(* Logix 5000 project; controller R400_500_XLS vendor 1 type 14 code 216 rev 31.11; software revision 31.01; part 26 of 32 *)
(* tags used below, declared in another part *)
   Abort1 : DINT;   // Not Used
   Alarm : SINT;   // Wait 3 seconds
   AlarmAcked : BOOL;   // Alarm has been acked
   bAlrm : BOOL[64];
   Chem_Pump : UDT_CHEM_PUMP[4];   // Chemical Pump flow rate
   ChemPumpIndex : DINT;
   CycExcBuffer : UDT_CYCLE;
   CycleSequence : UDT_CYCLE_SEQUENCE;
   Delta_T : REAL;
   DRYING : DINT;   // Drying id number
   F1rinse : DINT;   // Not Used
   F2rinse : DINT;   // Not Used
   F3rinse : DINT;   // Not Used
   FC22_SumpWaterVolume : REAL;   // Water volume
   FC22_Tran1 : BOOL;   // First transition
   FC22_Tran3 : BOOL;   // Third transition
   FC22_Tran4 : BOOL;   // Fourth transition
   FC22_WashIndex : SINT;
   HeatSmp : DINT;
   HighLimt : REAL;
   I_Pw_Tnk_Lvl_Sw_Deb : BOOL;   // Debounced pure water tank level switch (100ms)
   Inj_Time : SINT;   // Time based chemical injection steps
   LowLimt : REAL;
   M : DINT[5];   // Memory Bits
   MaxPressRecord : REAL;
   MinPressRecord : REAL;
   Neutral : SINT;
   ONS_FC17_1 : BOOL;
   ONS_FC17_2 : BOOL;
   ONS_FC22 : SINT;
   ONS_FC40 : SINT;
   ONS_WSH30 : SINT;
   PrintPressureDelay : DINT;
   PumpLowFRinse : DINT;   // Delay for pump low speed during final rinse treatment
   PumpLowPW_W_R : DINT;   // Delay for pump low speed during pre-wash, wash and rinse treatments
   PURE_WATER_HEATING_TIME : DINT;   // Time before an alarm is thrown when the pure water tank is heating
   PureWaterTankFilling : BOOL;   // Start PWT filling
   PW_HeatSp_5 : REAL;
   PW_HeatSp_X : REAL;
   PWHeat : SINT;
   Run : DINT;
   Service : DINT[2];   // Unused Service Mode Memory Bit
   StartPump1 : BOOL;   // Pump Low Speed
   StartPump2 : BOOL;   // Pump High Speed
   StartPump3 : BOOL;   // Main Pump running
   SUMP_HIGH_VOLUME_400 : REAL;   // High sump volume
   SUMP_HIGH_VOLUME_500 : REAL;
   SUMP_LOW_VOLUME_400 : REAL;   // Low sump volume
   SUMP_LOW_VOLUME_500 : REAL;
   SumpWaterVolume : DINT;   // Sump Water Volume 0 =Low 1= High
   T0_Temp : REAL;
   T1_Temp : REAL;
   TempChange : BOOL;
   Tmr : TIMER[107];
   Trt_PrWsh : DINT;
   Trt_Rinse : DINT;   // Rinse steps
   Trt_Wsh : DINT;
   WASH_1 : DINT;   // Wash 1 id number
   WASH_5 : DINT;   // Wash 5 id number
   WSH56_StartPump : BOOL;   // Start pump signal
   bPureWaterFillingAuthorization : BOOL;   // Pure Water Filling Authorization Signal
   I_Chm_1_Lvl_Sw : BOOL;   // Chemical Pump #1 level switch
   I_Chm_2_Lvl_Sw : BOOL;   // Chemical Pump #2 level switch
   I_Chm_3_Lvl_Sw : BOOL;   // Chemical Pump #3 level switch
   I_Chm_4_Lvl_Sw : BOOL;   // Chemical Pump #4 level switch
   I_MCR : BOOL;   // MCR input
   I_Mtr_Ovrld : BOOL;   // Motor overload
   I_Shlf_Sw : BOOL;   // Shelf switch
   PmpPres : REAL;
   PureWaterTankDrainingDeadLeg : BOOL;
   PureWaterTankFillingRequest : BOOL;
   PureWaterTankTemp : REAL;   // Pure water tank temperature
   Q_Pw_Tnk_Stm_Vlve : BOOL;   // PWT Steam Valve / Electric Heater
   SPV_19 : BOOL;   // Screen 80 Enabled/Disabled Pump pressure monitoring
   tDelayBeforeTankFillingAuthAlarm : TIMER;
   Tpb : DINT[11];
   tPureWaterTankClosingDelay : TIMER;
   TreatmentPtr : DINT;
   Unit : Hrdwre;   // Unit Configuration
(* MainProgram, continued *)

ROUTINE WSH_27_WSH_28_PURE_WATER_TANK   (* ladder *)
// This routine manages the filling, the draining and the heating of the pure water tank
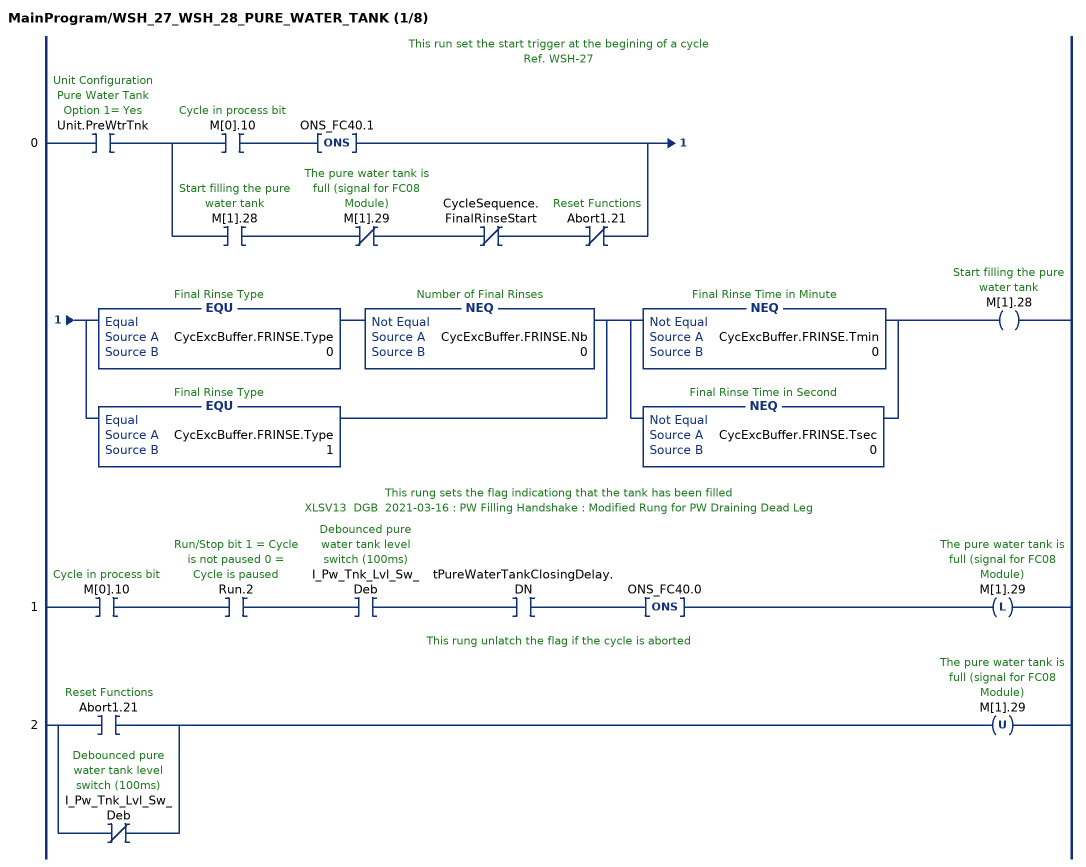
   // This run set the start trigger at the begining of a cycle
   // Ref. WSH-27
   0: XIC(Unit.PreWtrTnk)[XIC(M[0].10) ONS(ONS_FC40.1) ,XIC(M[1].28) XIO(M[1].29) XIO(CycleSequence.FinalRinseStart) XIO(Abort1.21) ][EQU(CycExcBuffer.FRINSE.Type,0) NEQ(CycExcBuffer.FRINSE.Nb,0) ,EQU(CycExcBuffer.FRINSE.Type,1) ][NEQ(CycExcBuffer.FRINSE.Tmin,0) ,NEQ(CycExcBuffer.FRINSE.Tsec,0) ]OTE(M[1].28);
   // This rung sets the flag indicationg that the tank has been filled
   // XLSV13  DGB  2021-03-16 : PW Filling Handshake : Modified Rung for PW Draining Dead Leg
   1: XIC(M[0].10)XIC(Run.2)XIC(I_Pw_Tnk_Lvl_Sw_Deb)XIC(tPureWaterTankClosingDelay.DN)ONS(ONS_FC40.0)OTL(M[1].29);
   // This rung unlatch the flag if the cycle is aborted
   2: [XIC(Abort1.21) ,XIO(I_Pw_Tnk_Lvl_Sw_Deb) ]OTU(M[1].29);
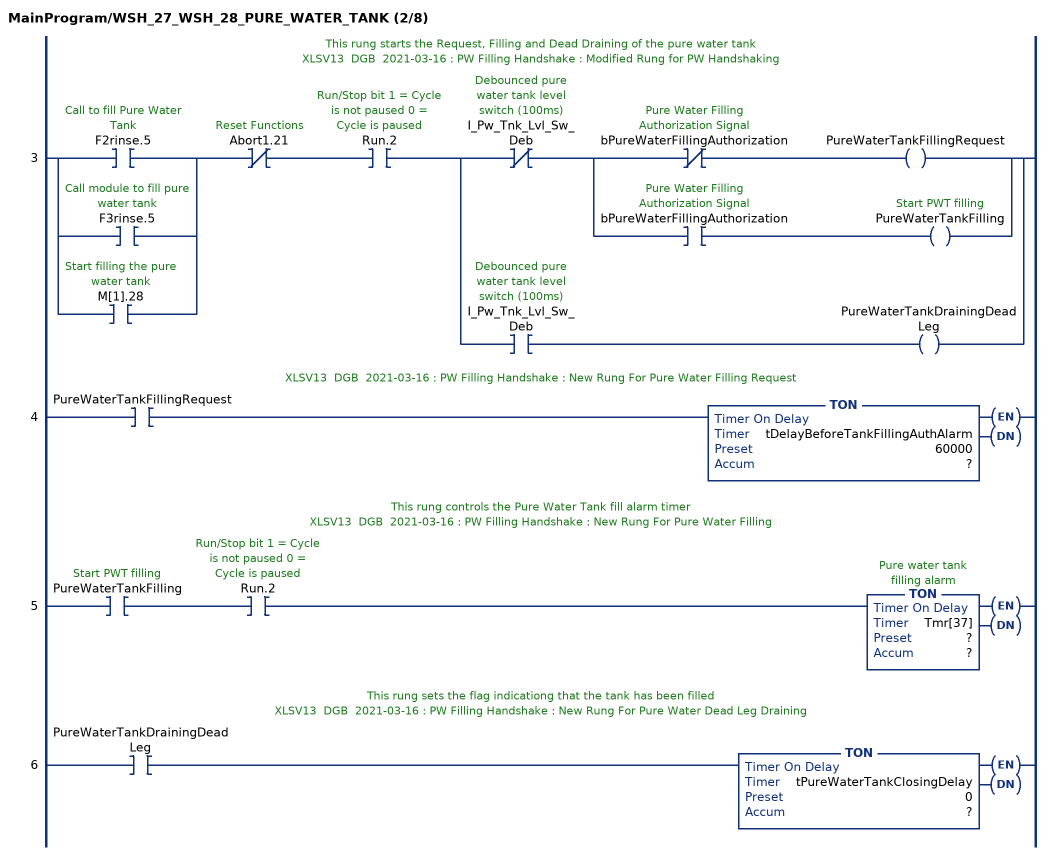
   // This rung starts the Request, Filling and Dead Draining of the pure water tank
   // XLSV13  DGB  2021-03-16 : PW Filling Handshake : Modified Rung for PW Handshaking
   3: [XIC(F2rinse.5) ,XIC(F3rinse.5) ,XIC(M[1].28) ]XIO(Abort1.21)XIC(Run.2)[XIO(I_Pw_Tnk_Lvl_Sw_Deb) [XIO(bPureWaterFillingAuthorization) OTE(PureWaterTankFillingRequest) ,XIC(bPureWaterFillingAuthorization) OTE(PureWaterTankFilling) ] ,XIC(I_Pw_Tnk_Lvl_Sw_Deb) OTE(PureWaterTankDrainingDeadLeg) ];
   // XLSV13  DGB  2021-03-16 : PW Filling Handshake : New Rung For Pure Water Filling Request
   4: XIC(PureWaterTankFillingRequest)TON(tDelayBeforeTankFillingAuthAlarm,?,?);
   // This rung controls the Pure Water Tank fill alarm timer
   // XLSV13  DGB  2021-03-16 : PW Filling Handshake : New Rung For Pure Water Filling
   5: XIC(PureWaterTankFilling)XIC(Run.2)TON(Tmr[37],?,?);
   // This rung sets the flag indicationg that the tank has been filled
   // XLSV13  DGB  2021-03-16 : PW Filling Handshake : New Rung For Pure Water Dead Leg Draining
   6: XIC(PureWaterTankDrainingDeadLeg)TON(tPureWaterTankClosingDelay,?,?);
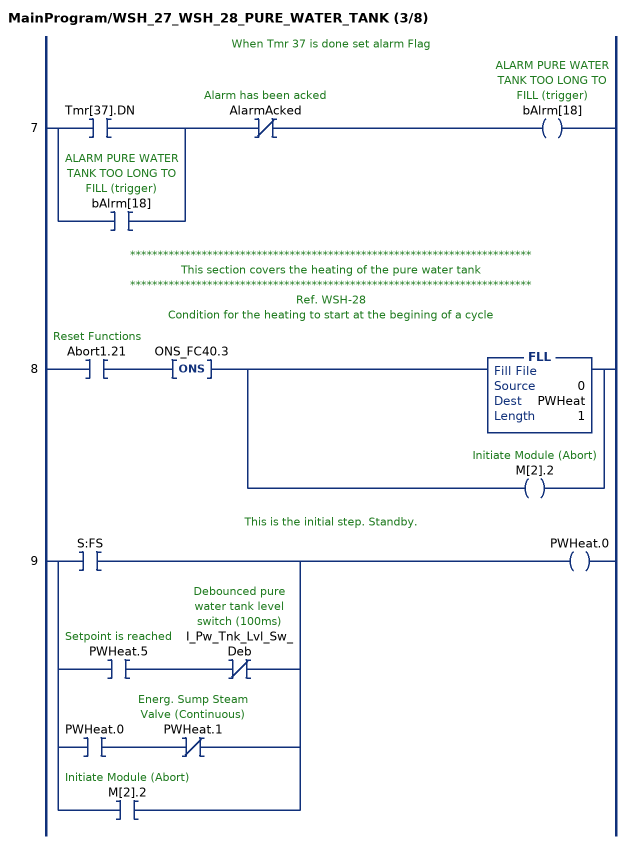
   // When Tmr 37 is done set alarm Flag
   7: [XIC(Tmr[37].DN) ,XIC(bAlrm[18]) ]XIO(AlarmAcked)OTE(bAlrm[18]);
   // *************************************************************************
   // This section covers the heating of the pure water tank
   // *************************************************************************
   // Ref. WSH-28
   // Condition for the heating to start at the begining of a cycle
   8: XIC(Abort1.21)ONS(ONS_FC40.3)[FLL(0,PWHeat,1) ,OTE(M[2].2) ];
   // This is the initial step. Standby.
   9: [XIC(S:FS) ,XIC(PWHeat.5) XIO(I_Pw_Tnk_Lvl_Sw_Deb) ,XIC(PWHeat.0) XIO(PWHeat.1) ,XIC(M[2].2) ]OTE(PWHeat.0);
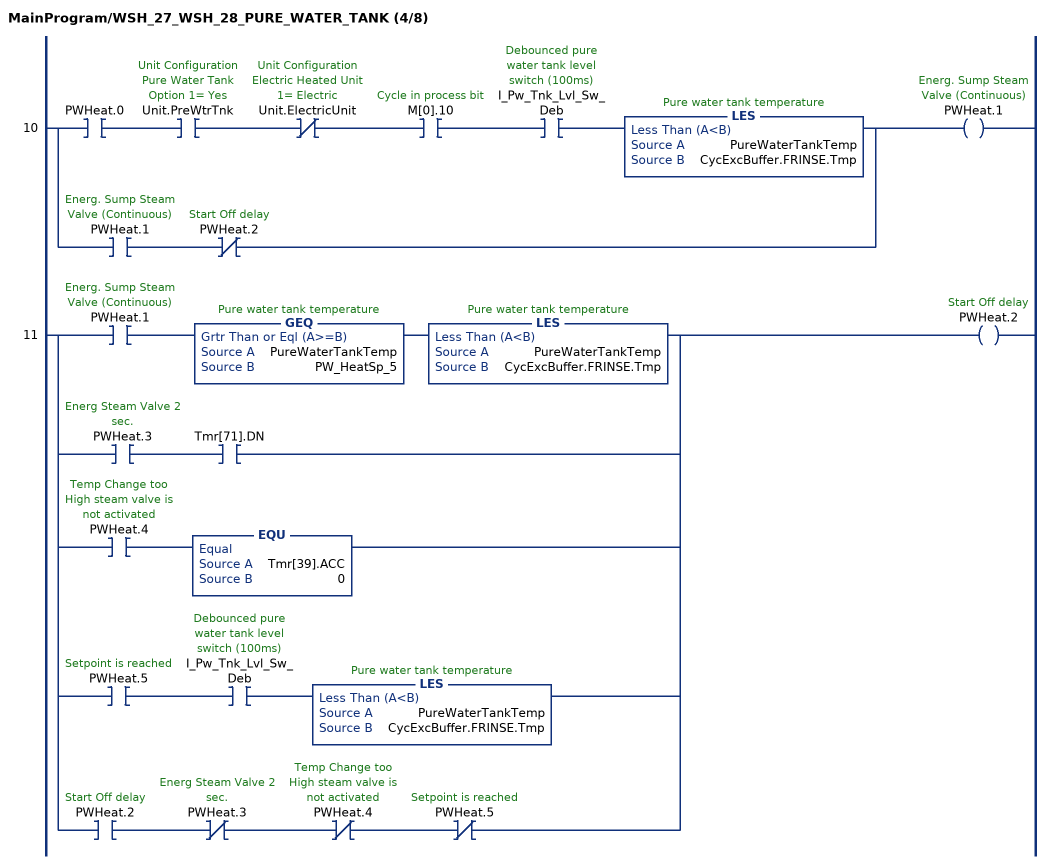
   10: [XIC(PWHeat.0) XIC(Unit.PreWtrTnk) XIO(Unit.ElectricUnit) XIC(M[0].10) XIC(I_Pw_Tnk_Lvl_Sw_Deb) LES(PureWaterTankTemp,CycExcBuffer.FRINSE.Tmp) ,XIC(PWHeat.1) XIO(PWHeat.2) ]OTE(PWHeat.1);
   11: [XIC(PWHeat.1) GEQ(PureWaterTankTemp,PW_HeatSp_5) LES(PureWaterTankTemp,CycExcBuffer.FRINSE.Tmp) ,XIC(PWHeat.3) XIC(Tmr[71].DN) ,XIC(PWHeat.4) EQU(Tmr[39].ACC,0) ,XIC(PWHeat.5) XIC(I_Pw_Tnk_Lvl_Sw_Deb) LES(PureWaterTankTemp,CycExcBuffer.FRINSE.Tmp) ,XIC(PWHeat.2) XIO(PWHeat.3) XIO(PWHeat.4) XIO(PWHeat.5) ]OTE(PWHeat.2);
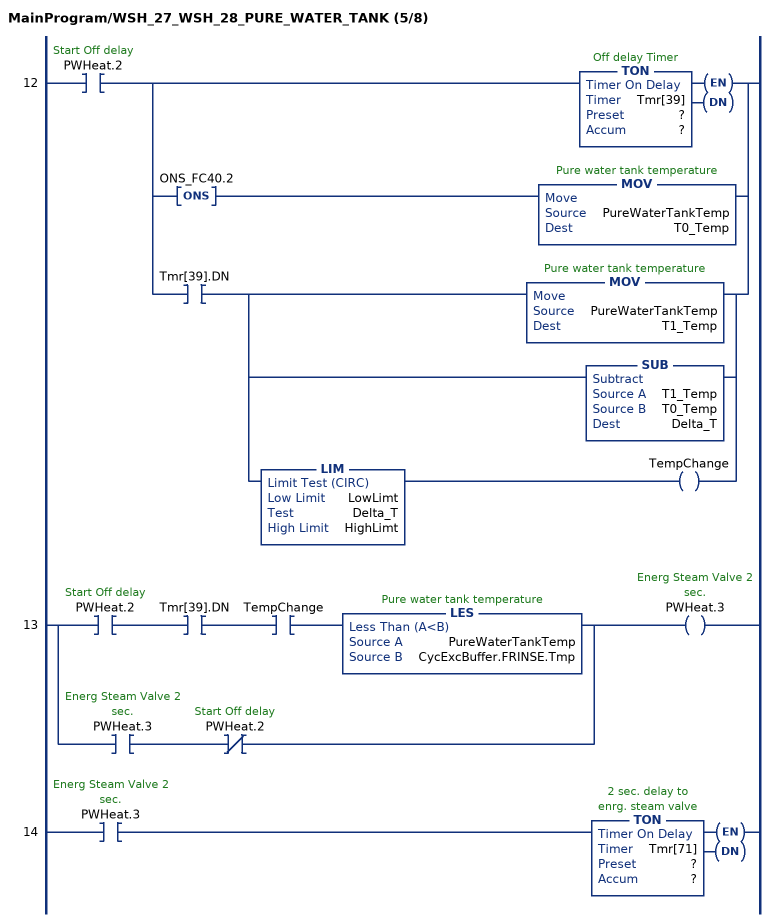
   12: XIC(PWHeat.2)[TON(Tmr[39],?,?) ,ONS(ONS_FC40.2) MOV(PureWaterTankTemp,T0_Temp) ,XIC(Tmr[39].DN) [MOV(PureWaterTankTemp,T1_Temp) ,SUB(T1_Temp,T0_Temp,Delta_T) ,LIM(LowLimt,Delta_T,HighLimt) OTE(TempChange) ] ];
   13: [XIC(PWHeat.2) XIC(Tmr[39].DN) XIC(TempChange) LES(PureWaterTankTemp,CycExcBuffer.FRINSE.Tmp) ,XIC(PWHeat.3) XIO(PWHeat.2) ]OTE(PWHeat.3);
   14: XIC(PWHeat.3)TON(Tmr[71],?,?);
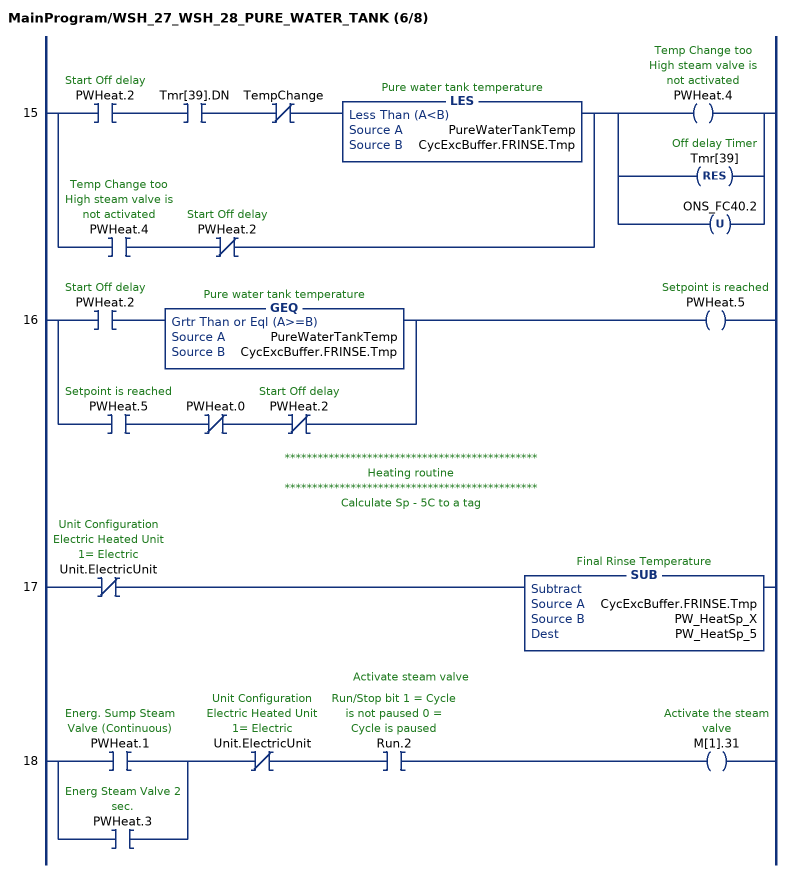
   15: [XIC(PWHeat.2) XIC(Tmr[39].DN) XIO(TempChange) LES(PureWaterTankTemp,CycExcBuffer.FRINSE.Tmp) ,XIC(PWHeat.4) XIO(PWHeat.2) ][OTE(PWHeat.4) ,RES(Tmr[39]) ,OTU(ONS_FC40.2) ];
   16: [XIC(PWHeat.2) GEQ(PureWaterTankTemp,CycExcBuffer.FRINSE.Tmp) ,XIC(PWHeat.5) XIO(PWHeat.0) XIO(PWHeat.2) ]OTE(PWHeat.5);
   // **********************************************
   // Heating routine
   // **********************************************
   // Calculate Sp - 5C to a tag
   17: XIO(Unit.ElectricUnit)SUB(CycExcBuffer.FRINSE.Tmp,PW_HeatSp_X,PW_HeatSp_5);
   // Activate steam valve
   18: [XIC(PWHeat.1) ,XIC(PWHeat.3) ]XIO(Unit.ElectricUnit)XIC(Run.2)OTE(M[1].31);
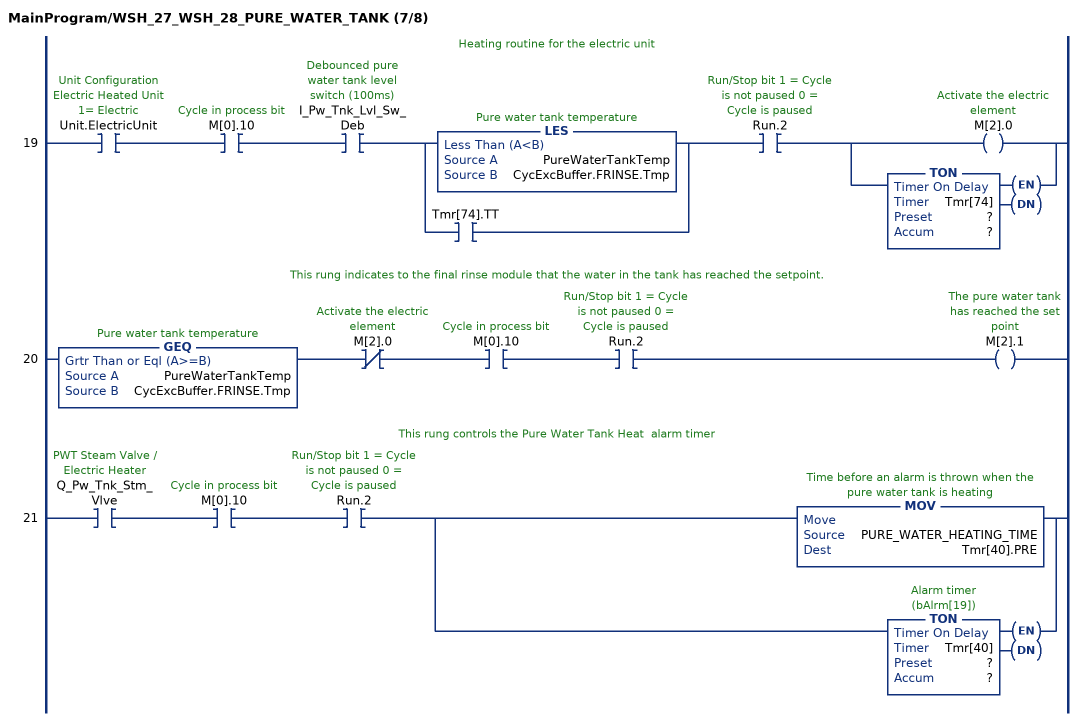
   // Heating routine for the electric unit
   19: XIC(Unit.ElectricUnit)XIC(M[0].10)XIC(I_Pw_Tnk_Lvl_Sw_Deb)[LES(PureWaterTankTemp,CycExcBuffer.FRINSE.Tmp) ,XIC(Tmr[74].TT) ]XIC(Run.2)[OTE(M[2].0) ,TON(Tmr[74],?,?) ];
   // This rung indicates to the final rinse module that the water in the tank has reached the setpoint.
   20: GEQ(PureWaterTankTemp,CycExcBuffer.FRINSE.Tmp)XIO(M[2].0)XIC(M[0].10)XIC(Run.2)OTE(M[2].1);
   // This rung controls the Pure Water Tank Heat  alarm timer
   21: XIC(Q_Pw_Tnk_Stm_Vlve)XIC(M[0].10)XIC(Run.2)[MOV(PURE_WATER_HEATING_TIME,Tmr[40].PRE) ,TON(Tmr[40],?,?) ];
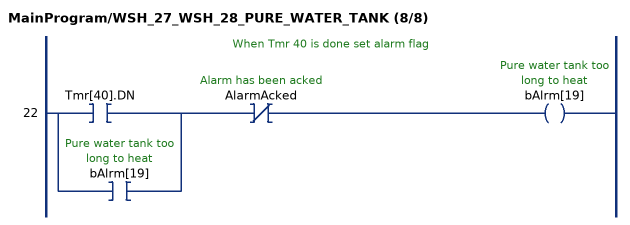
   // When Tmr 40 is done set alarm flag
   22: [XIC(Tmr[40].DN) ,XIC(bAlrm[19]) ]XIO(AlarmAcked)OTE(bAlrm[19]);
END_ROUTINE

ROUTINE WSH_29_START_PUMP   (* ladder *)
// This module starts the main pump
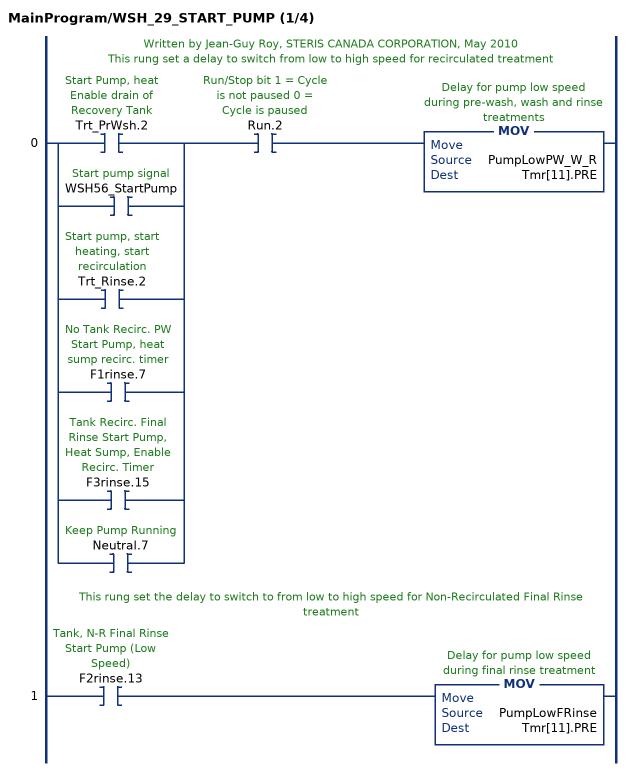
   // Written by Jean-Guy Roy, STERIS CANADA CORPORATION, May 2010
   // This rung set a delay to switch from low to high speed for recirculated treatment
   0: [XIC(Trt_PrWsh.2) ,XIC(WSH56_StartPump) ,XIC(Trt_Rinse.2) ,XIC(F1rinse.7) ,XIC(F3rinse.15) ,XIC(Neutral.7) ]XIC(Run.2)MOV(PumpLowPW_W_R,Tmr[11].PRE);
   // This rung set the delay to switch to from low to high speed for Non-Recirculated Final Rinse treatment
   1: XIC(F2rinse.13)MOV(PumpLowFRinse,Tmr[11].PRE);
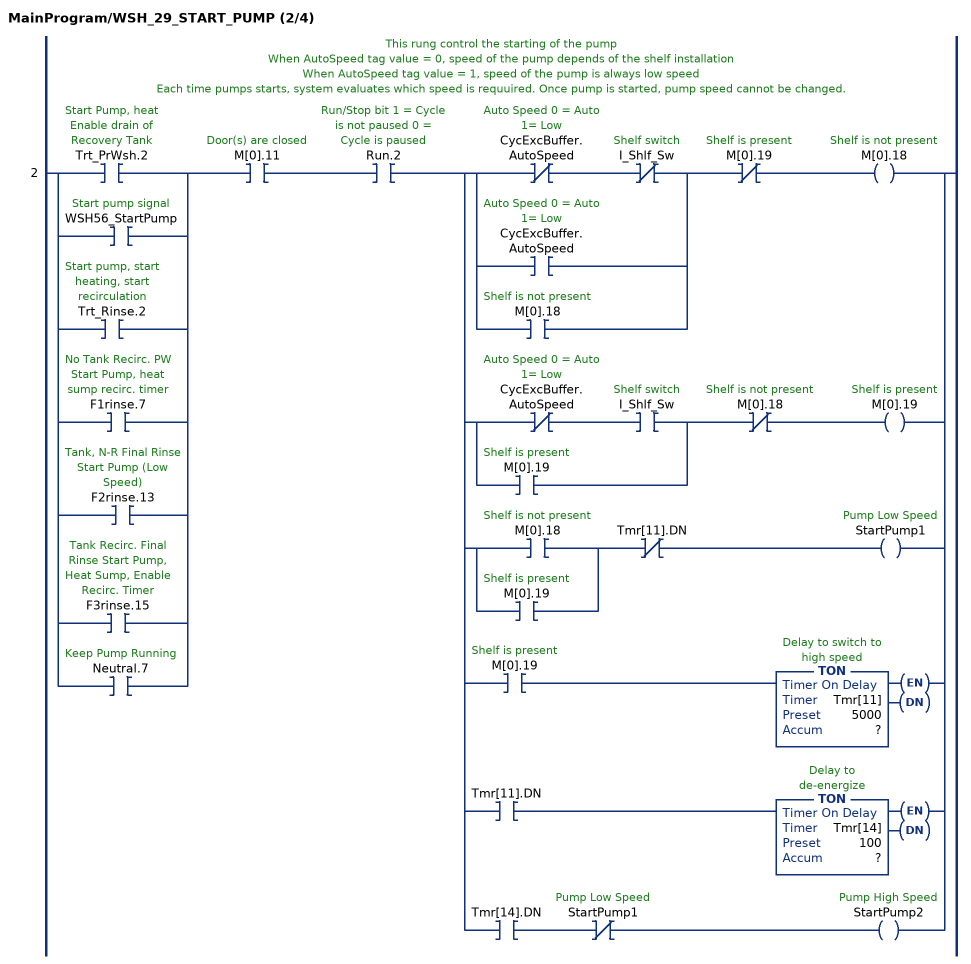
   // This rung control the starting of the pump
   // When AutoSpeed tag value = 0, speed of the pump depends of the shelf installation
   // When AutoSpeed tag value = 1, speed of the pump is always low speed
   // Each time pumps starts, system evaluates which speed is requuired. Once pump is started, pump speed cannot be changed.
   2: [XIC(Trt_PrWsh.2) ,XIC(WSH56_StartPump) ,XIC(Trt_Rinse.2) ,XIC(F1rinse.7) ,XIC(F2rinse.13) ,XIC(F3rinse.15) ,XIC(Neutral.7) ]XIC(M[0].11)XIC(Run.2)[[XIO(CycExcBuffer.AutoSpeed) XIO(I_Shlf_Sw) ,XIC(CycExcBuffer.AutoSpeed) ,XIC(M[0].18) ] XIO(M[0].19) OTE(M[0].18) ,[XIO(CycExcBuffer.AutoSpeed) XIC(I_Shlf_Sw) ,XIC(M[0].19) ] XIO(M[0].18) OTE(M[0].19) ,[XIC(M[0].18) ,XIC(M[0].19) ] XIO(Tmr[11].DN) OTE(StartPump1) ,XIC(M[0].19) TON(Tmr[11],?,?) ,XIC(Tmr[11].DN) TON(Tmr[14],?,?) ,XIC(Tmr[14].DN) XIO(StartPump1) OTE(StartPump2) ];
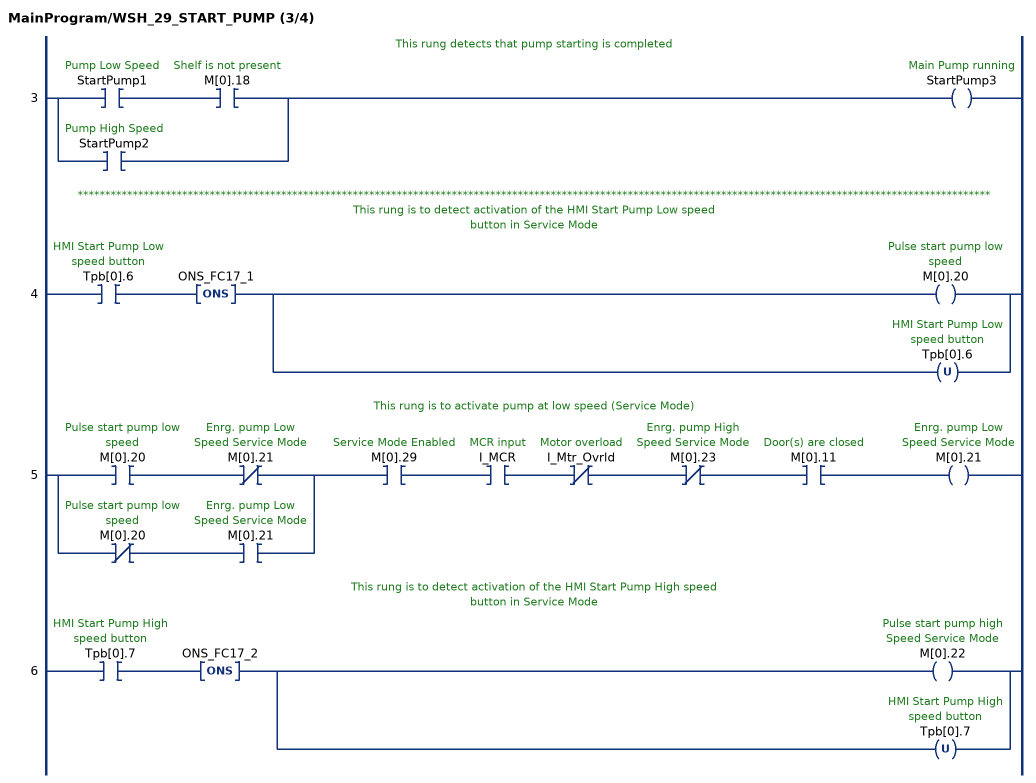
   // This rung detects that pump starting is completed
   3: [XIC(StartPump1) XIC(M[0].18) ,XIC(StartPump2) ]OTE(StartPump3);
   // **********************************************************************************************************************************************************************
   // This rung is to detect activation of the HMI Start Pump Low speed
   // button in Service Mode
   4: XIC(Tpb[0].6)ONS(ONS_FC17_1)[OTE(M[0].20) ,OTU(Tpb[0].6) ];
   // This rung is to activate pump at low speed (Service Mode)
   5: [XIC(M[0].20) XIO(M[0].21) ,XIO(M[0].20) XIC(M[0].21) ]XIC(M[0].29)XIC(I_MCR)XIO(I_Mtr_Ovrld)XIO(M[0].23)XIC(M[0].11)OTE(M[0].21);
   // This rung is to detect activation of the HMI Start Pump High speed
   // button in Service Mode
   6: XIC(Tpb[0].7)ONS(ONS_FC17_2)[OTE(M[0].22) ,OTU(Tpb[0].7) ];
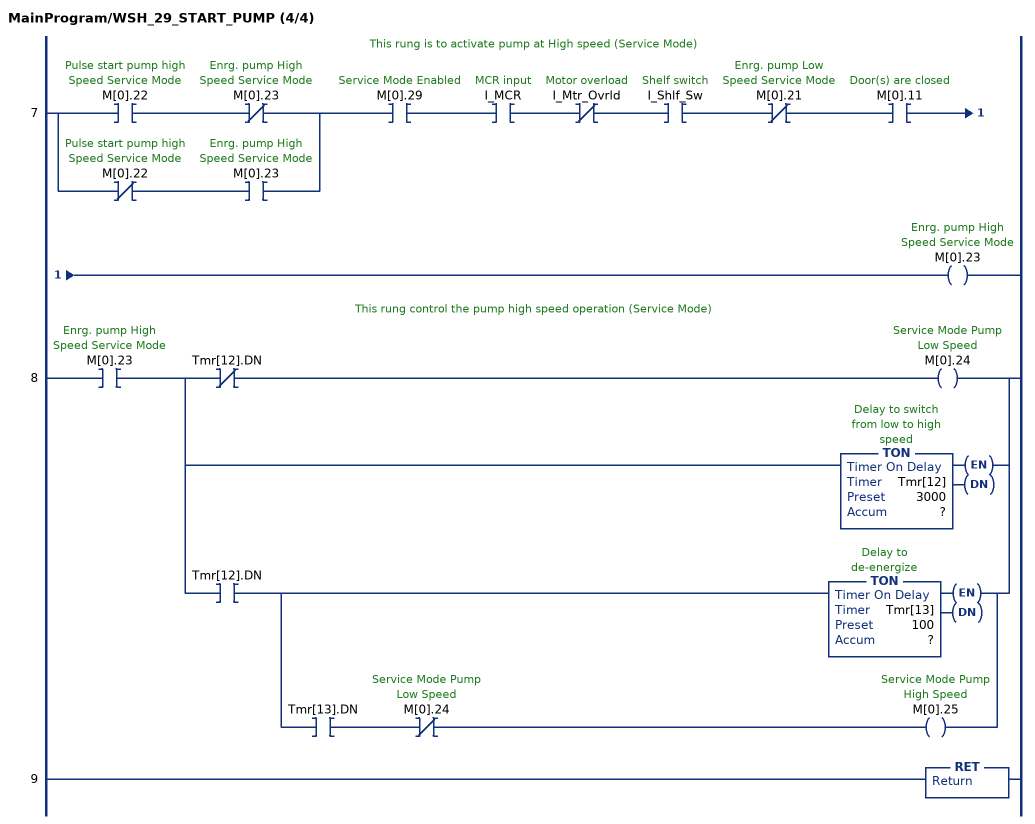
   // This rung is to activate pump at High speed (Service Mode)
   7: [XIC(M[0].22) XIO(M[0].23) ,XIO(M[0].22) XIC(M[0].23) ]XIC(M[0].29)XIC(I_MCR)XIO(I_Mtr_Ovrld)XIC(I_Shlf_Sw)XIO(M[0].21)XIC(M[0].11)OTE(M[0].23);
   // This rung control the pump high speed operation (Service Mode)
   8: XIC(M[0].23)[XIO(Tmr[12].DN) OTE(M[0].24) ,TON(Tmr[12],?,?) ,XIC(Tmr[12].DN) [TON(Tmr[13],?,?) ,XIC(Tmr[13].DN) XIO(M[0].24) OTE(M[0].25) ] ];
   9: RET();
END_ROUTINE

ROUTINE WSH_30_MONITOR_PRESSURE   (* ladder *)
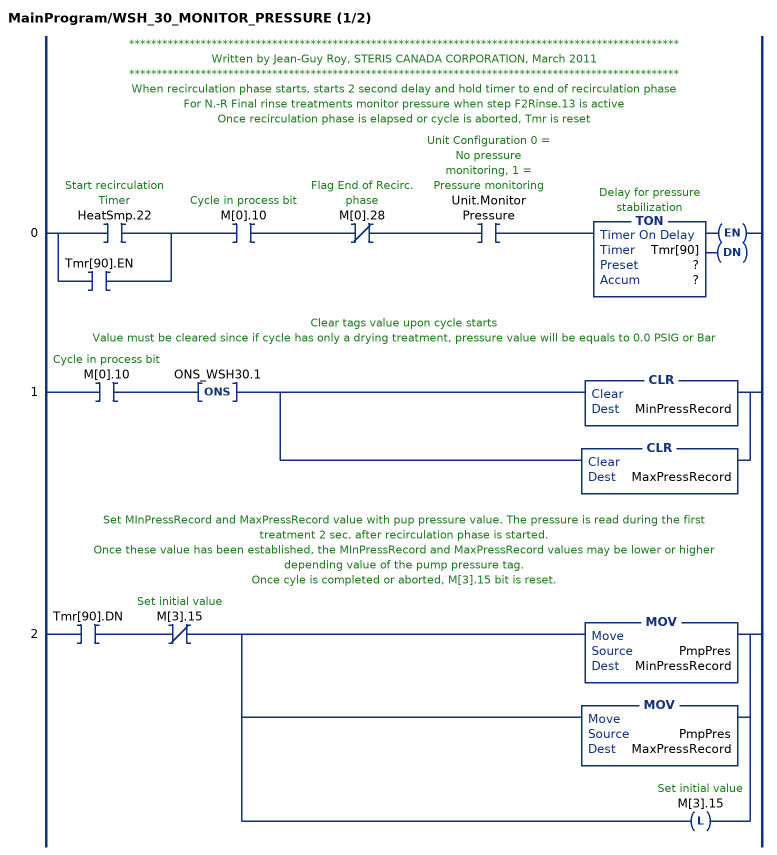
   // ****************************************************************************************************
   // Written by Jean-Guy Roy, STERIS CANADA CORPORATION, March 2011
   // ****************************************************************************************************
   // When recirculation phase starts, starts 2 second delay and hold timer to end of recirculation phase
   // For N.-R Final rinse treatments monitor pressure when step F2Rinse.13 is active
   // Once recirculation phase is elapsed or cycle is aborted, Tmr is reset
   0: [XIC(HeatSmp.22) ,XIC(Tmr[90].EN) ]XIC(M[0].10)XIO(M[0].28)XIC(Unit.MonitorPressure)TON(Tmr[90],?,?);
   // Clear tags value upon cycle starts
   // Value must be cleared since if cycle has only a drying treatment, pressure value will be equals to 0.0 PSIG or Bar
   1: XIC(M[0].10)ONS(ONS_WSH30.1)[CLR(MinPressRecord) ,CLR(MaxPressRecord) ];
   // Set MInPressRecord and MaxPressRecord value with pup pressure value. The pressure is read during the first treatment 2 sec. after recirculation phase is started.
   // Once these value has been established, the MInPressRecord and MaxPressRecord values may be lower or higher depending value of the pump pressure tag.
   // Once cyle is completed or aborted, M[3].15 bit is reset.
   2: XIC(Tmr[90].DN)XIO(M[3].15)[MOV(PmpPres,MinPressRecord) ,MOV(PmpPres,MaxPressRecord) ,OTL(M[3].15) ];
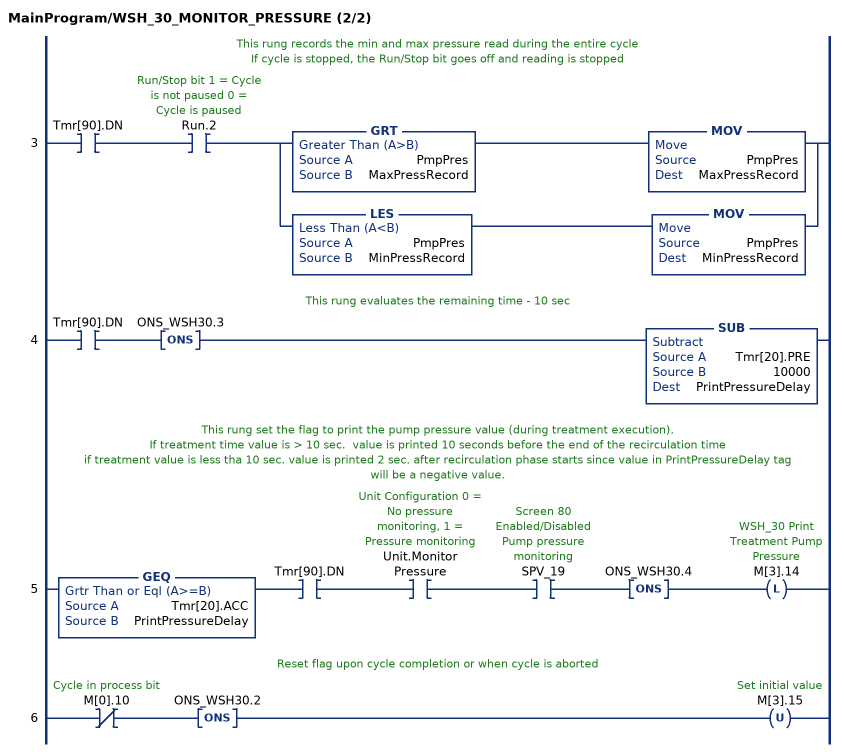
   // This rung records the min and max pressure read during the entire cycle
   // If cycle is stopped, the Run/Stop bit goes off and reading is stopped
   3: XIC(Tmr[90].DN)XIC(Run.2)[GRT(PmpPres,MaxPressRecord) MOV(PmpPres,MaxPressRecord) ,LES(PmpPres,MinPressRecord) MOV(PmpPres,MinPressRecord) ];
   // This rung evaluates the remaining time - 10 sec
   4: XIC(Tmr[90].DN)ONS(ONS_WSH30.3)SUB(Tmr[20].PRE,10000,PrintPressureDelay);
   // This rung set the flag to print the pump pressure value (during treatment execution).
   // If treatment time value is > 10 sec.  value is printed 10 seconds before the end of the recirculation time
   // if treatment value is less tha 10 sec. value is printed 2 sec. after recirculation phase starts since value in PrintPressureDelay tag will be a negative value.
   5: GEQ(Tmr[20].ACC,PrintPressureDelay)XIC(Tmr[90].DN)XIC(Unit.MonitorPressure)XIC(SPV_19)ONS(ONS_WSH30.4)OTL(M[3].14);
   // Reset flag upon cycle completion or when cycle is aborted
   6: XIO(M[0].10)ONS(ONS_WSH30.2)OTU(M[3].15);
END_ROUTINE

ROUTINE WSH_32_TIME_BASED_INJECTION   (* ladder *)
// This routine manages the time based chemical injection
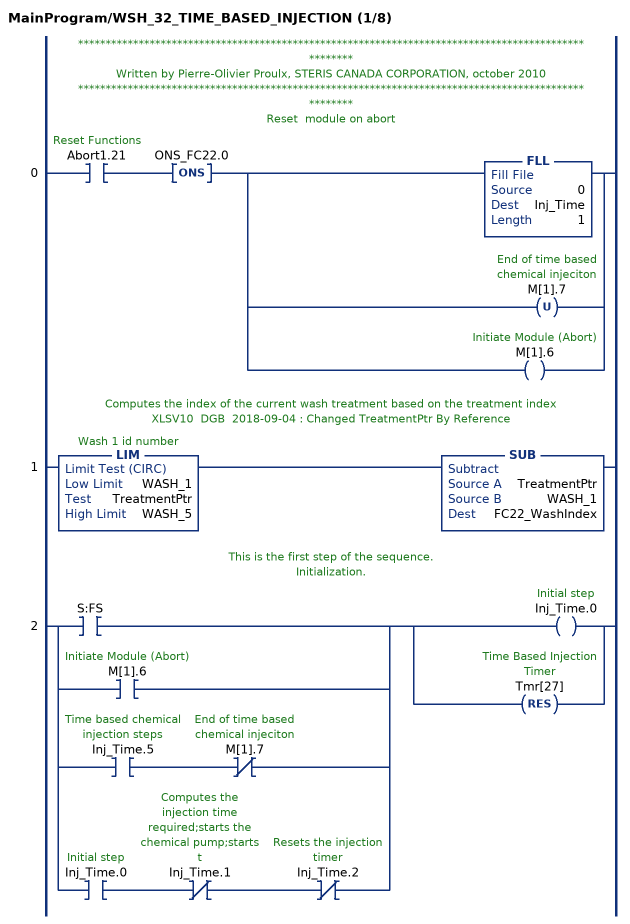
   // ****************************************************************************************************
   // Written by Pierre-Olivier Proulx, STERIS CANADA CORPORATION, october 2010
   // ****************************************************************************************************
   // Reset  module on abort
   0: XIC(Abort1.21)ONS(ONS_FC22.0)[FLL(0,Inj_Time,1) ,OTU(M[1].7) ,OTE(M[1].6) ];
   // Computes the index of the current wash treatment based on the treatment index
   // XLSV10  DGB  2018-09-04 : Changed TreatmentPtr By Reference
   1: LIM(WASH_1,TreatmentPtr,WASH_5)SUB(TreatmentPtr,WASH_1,FC22_WashIndex);
   // This is the first step of the sequence.
   // Initialization.
   2: [XIC(S:FS) ,XIC(M[1].6) ,XIC(Inj_Time.5) XIO(M[1].7) ,XIC(Inj_Time.0) XIO(Inj_Time.1) XIO(Inj_Time.2) ][OTE(Inj_Time.0) ,RES(Tmr[27]) ];
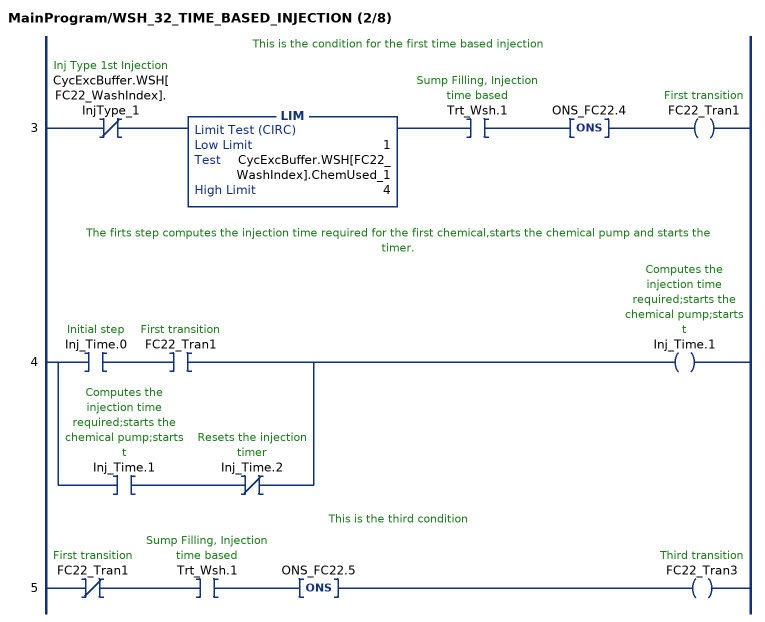
   // This is the condition for the first time based injection
   3: XIO(CycExcBuffer.WSH[FC22_WashIndex].InjType_1)LIM(1,CycExcBuffer.WSH[FC22_WashIndex].ChemUsed_1,4)XIC(Trt_Wsh.1)ONS(ONS_FC22.4)OTE(FC22_Tran1);
   // The firts step computes the injection time required for the first chemical,starts the chemical pump and starts the timer.
   4: [XIC(Inj_Time.0) XIC(FC22_Tran1) ,XIC(Inj_Time.1) XIO(Inj_Time.2) ]OTE(Inj_Time.1);
   // This is the third condition
   5: XIO(FC22_Tran1)XIC(Trt_Wsh.1)ONS(ONS_FC22.5)OTE(FC22_Tran3);
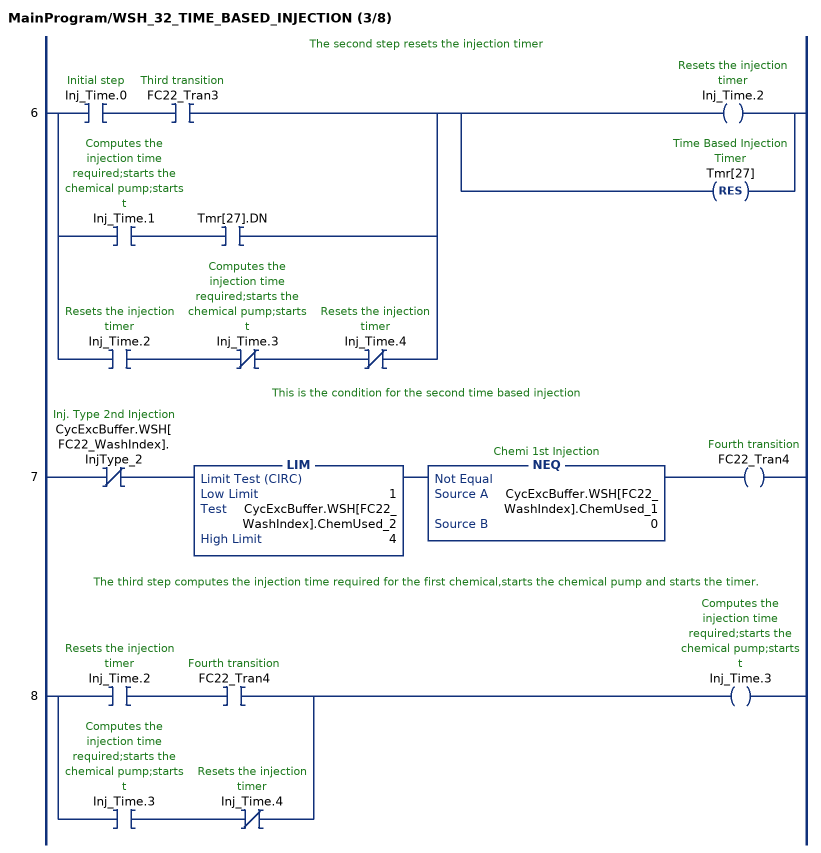
   // The second step resets the injection timer
   6: [XIC(Inj_Time.0) XIC(FC22_Tran3) ,XIC(Inj_Time.1) XIC(Tmr[27].DN) ,XIC(Inj_Time.2) XIO(Inj_Time.3) XIO(Inj_Time.4) ][OTE(Inj_Time.2) ,RES(Tmr[27]) ];
   // This is the condition for the second time based injection
   7: XIO(CycExcBuffer.WSH[FC22_WashIndex].InjType_2)LIM(1,CycExcBuffer.WSH[FC22_WashIndex].ChemUsed_2,4)NEQ(CycExcBuffer.WSH[FC22_WashIndex].ChemUsed_1,0)OTE(FC22_Tran4);
   // The third step computes the injection time required for the first chemical,starts the chemical pump and starts the timer.
   8: [XIC(Inj_Time.2) XIC(FC22_Tran4) ,XIC(Inj_Time.3) XIO(Inj_Time.4) ]OTE(Inj_Time.3);
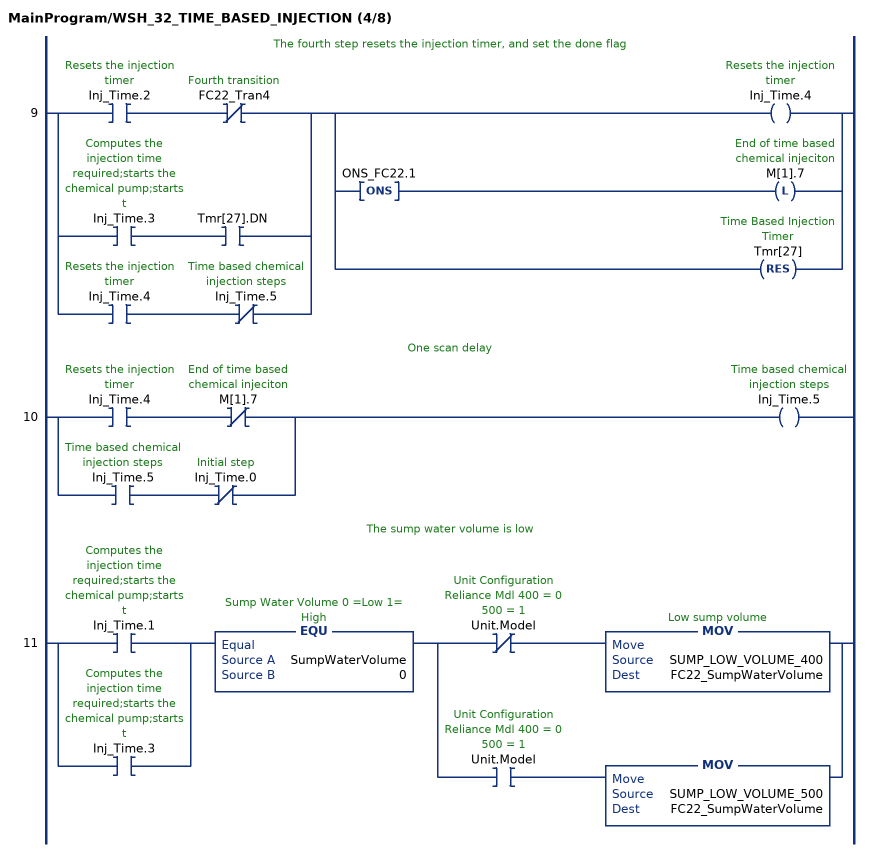
   // The fourth step resets the injection timer, and set the done flag
   9: [XIC(Inj_Time.2) XIO(FC22_Tran4) ,XIC(Inj_Time.3) XIC(Tmr[27].DN) ,XIC(Inj_Time.4) XIO(Inj_Time.5) ][OTE(Inj_Time.4) ,ONS(ONS_FC22.1) OTL(M[1].7) ,RES(Tmr[27]) ];
   // One scan delay
   10: [XIC(Inj_Time.4) XIO(M[1].7) ,XIC(Inj_Time.5) XIO(Inj_Time.0) ]OTE(Inj_Time.5);
   // The sump water volume is low
   11: [XIC(Inj_Time.1) ,XIC(Inj_Time.3) ]EQU(SumpWaterVolume,0)[XIO(Unit.Model) MOV(SUMP_LOW_VOLUME_400,FC22_SumpWaterVolume) ,XIC(Unit.Model) MOV(SUMP_LOW_VOLUME_500,FC22_SumpWaterVolume) ];
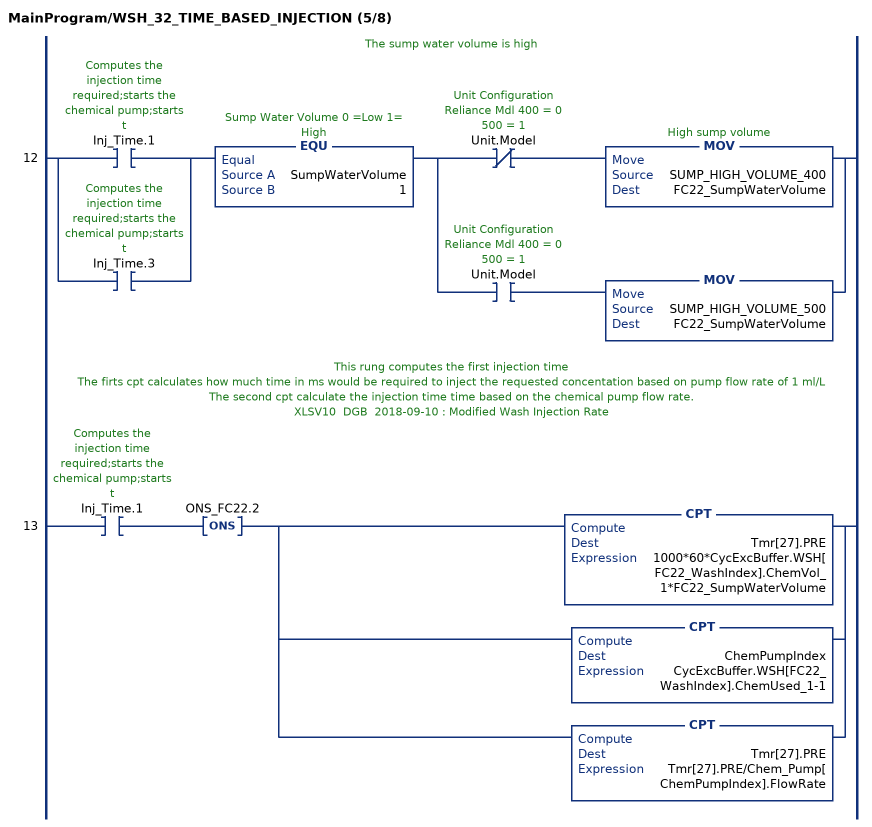
   // The sump water volume is high
   12: [XIC(Inj_Time.1) ,XIC(Inj_Time.3) ]EQU(SumpWaterVolume,1)[XIO(Unit.Model) MOV(SUMP_HIGH_VOLUME_400,FC22_SumpWaterVolume) ,XIC(Unit.Model) MOV(SUMP_HIGH_VOLUME_500,FC22_SumpWaterVolume) ];
   // This rung computes the first injection time
   // The firts cpt calculates how much time in ms would be required to inject the requested concentation based on pump flow rate of 1 ml/L
   // The second cpt calculate the injection time time based on the chemical pump flow rate.
   // XLSV10  DGB  2018-09-10 : Modified Wash Injection Rate
   13: XIC(Inj_Time.1)ONS(ONS_FC22.2)[CPT(Tmr[27].PRE,1000*60*CycExcBuffer.WSH[FC22_WashIndex].ChemVol_1*FC22_SumpWaterVolume) ,CPT(ChemPumpIndex,CycExcBuffer.WSH[FC22_WashIndex].ChemUsed_1-1) ,CPT(Tmr[27].PRE,Tmr[27].PRE/Chem_Pump[ChemPumpIndex].FlowRate) ];
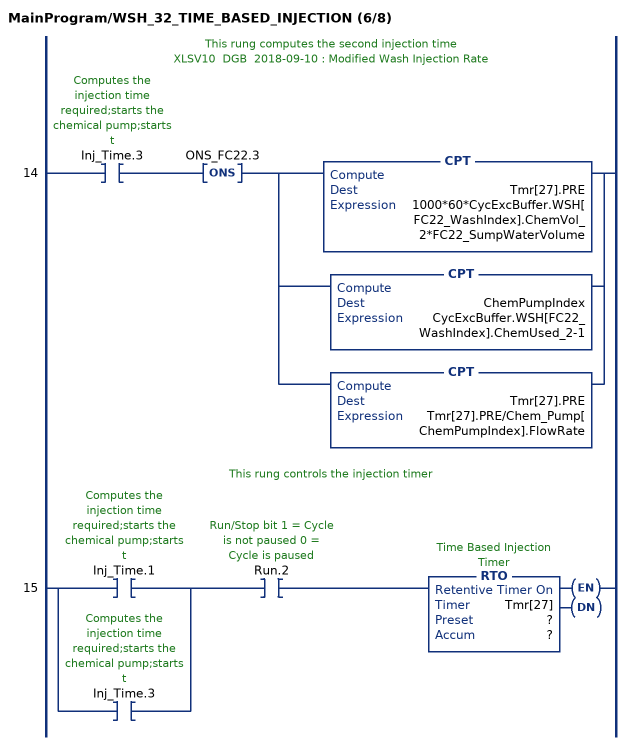
   // This rung computes the second injection time
   // XLSV10  DGB  2018-09-10 : Modified Wash Injection Rate
   14: XIC(Inj_Time.3)ONS(ONS_FC22.3)[CPT(Tmr[27].PRE,1000*60*CycExcBuffer.WSH[FC22_WashIndex].ChemVol_2*FC22_SumpWaterVolume) ,CPT(ChemPumpIndex,CycExcBuffer.WSH[FC22_WashIndex].ChemUsed_2-1) ,CPT(Tmr[27].PRE,Tmr[27].PRE/Chem_Pump[ChemPumpIndex].FlowRate) ];
   // This rung controls the injection timer
   15: [XIC(Inj_Time.1) ,XIC(Inj_Time.3) ]XIC(Run.2)RTO(Tmr[27],?,?);
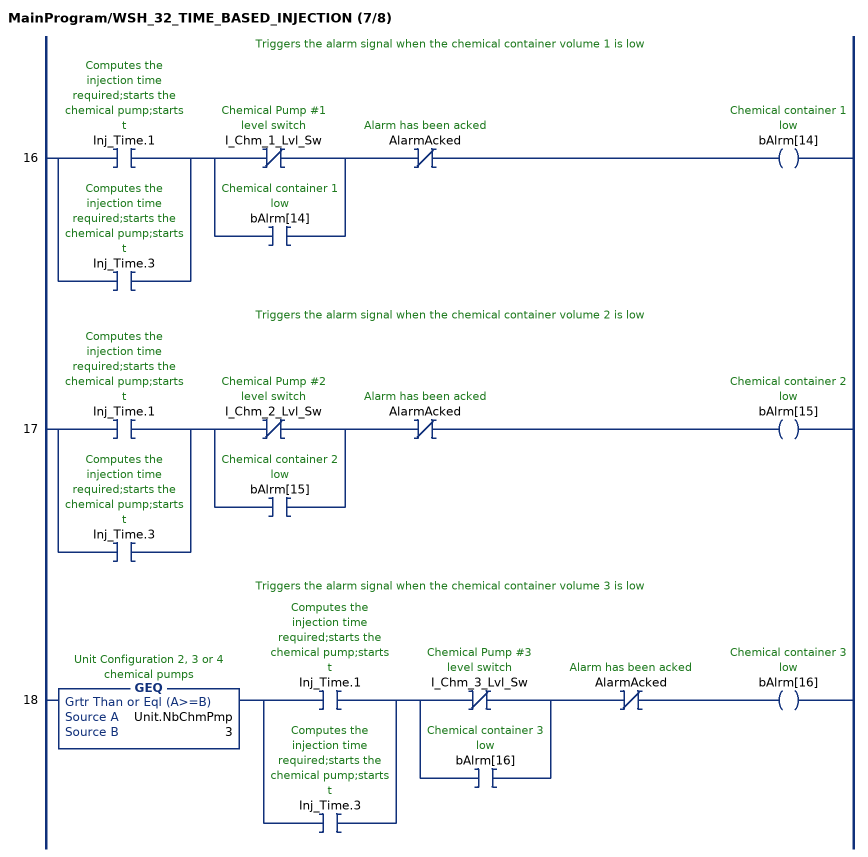
   // Triggers the alarm signal when the chemical container volume 1 is low
   16: [XIC(Inj_Time.1) ,XIC(Inj_Time.3) ][XIO(I_Chm_1_Lvl_Sw) ,XIC(bAlrm[14]) ]XIO(AlarmAcked)OTE(bAlrm[14]);
   // Triggers the alarm signal when the chemical container volume 2 is low
   17: [XIC(Inj_Time.1) ,XIC(Inj_Time.3) ][XIO(I_Chm_2_Lvl_Sw) ,XIC(bAlrm[15]) ]XIO(AlarmAcked)OTE(bAlrm[15]);
   // Triggers the alarm signal when the chemical container volume 3 is low
   18: GEQ(Unit.NbChmPmp,3)[XIC(Inj_Time.1) ,XIC(Inj_Time.3) ][XIO(I_Chm_3_Lvl_Sw) ,XIC(bAlrm[16]) ]XIO(AlarmAcked)OTE(bAlrm[16]);
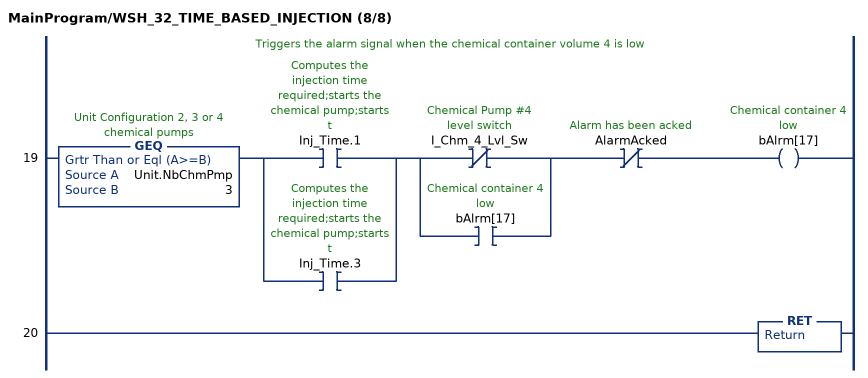
   // Triggers the alarm signal when the chemical container volume 4 is low
   19: GEQ(Unit.NbChmPmp,3)[XIC(Inj_Time.1) ,XIC(Inj_Time.3) ][XIO(I_Chm_4_Lvl_Sw) ,XIC(bAlrm[17]) ]XIO(AlarmAcked)OTE(bAlrm[17]);
   20: RET();
END_ROUTINE
